Fanuc KAREL source: kt00267.KL

-- PROVISIONAL review KL for V1013-1; original PC SHA256 f7ed19ebe923b0019c9fd7f40b6310b46c5a861f0aa85319aa3adadf6d86af20
-- Incomplete behavior may be omitted. Consult companion uncertainty JSON. Do not deploy.
PROGRAM KT00267
%NOLOCKGROUP
VAR
  I2 : INTEGER
  OUT : BOOLEAN
-- UNRESOLVED_DECL Y1 type=002018
BEGIN
  -- UNRESOLVED_PC offsets 5-19; opcodes 2E,22,9D,33,B2
  -- UNRESOLVED_PC offsets 24-35; opcodes 2E,23
  -- UNRESOLVED_PC offsets 40-62; opcodes 22,9D,33,B1,21,57,23
  -- UNRESOLVED_PC offsets 67-71; opcodes 7F
END KT00267
